TYPE E_WorkingMode :(	
	eManualMode			:=0,
	eSemiAutoMode		:=1,
	eAutoMode			:=2);
END_TYPE

//eWorkingModeNone	:=0,

(* stored: Version 1.1.0.1, ProductVersion 3.1.4024.13
   DUT E_WorkingMode: Id {5647a93a-b620-42e2-bf82-39ca71d039d4} *)
